// TwinCAT 3 PLC project Untitled1
// ProgramVersion: 3.1.4026.27
// libraries:
//   Tc2_Standard, * (Beckhoff Automation GmbH)
//   Tc2_System, * (Beckhoff Automation GmbH)
//   Tc3_EventLogger, * (Beckhoff Automation GmbH)
//   Tc3_Module, * (Beckhoff Automation GmbH)
//   VisuDialogs, * (System)
//   VisuSymbols,4.5.0.0,System
// project tree:
//   / GlobalTextList.TcGTLO, PlcTask.TcTTO, Visualization Manager.TcVMO (not stored)
//   GVLs/ gAL.TcGVL
//   POUs/Alarms_and_Emergency/ Alarm_System.TcPOU, FB_Emergency_Shutdown.TcPOU, FB_Alarm.TcPOU
//   POUs/ FB_ControlPanel.TcPOU, FB_Scale.TcPOU, MAIN.TcPOU, PI_Function_Block.TcPOU
// real-time tasks:
//   TASK PlcTask: cycle T#10ms, priority 20, ADS port 350
// I/O:
//   DEVICE Device 1 (EtherCAT), AmsNetId 10.0.0.14.2.1
//     Term 7 (EK1200) [EK1200-5000 EtherCAT Power supply (2A E-Bus)]
//       Term 2 (EL4004) [EL4004 4Ch. Ana. Output 0-10V, 12bit]
//       Term 3 (EL4004) [EL4004 4Ch. Ana. Output 0-10V, 12bit]
//       Term 8 (EL3024) [EL3024 4Ch. Ana. Input 4-20mA DIFF]
//       Term 9 (EL3024) [EL3024 4Ch. Ana. Input 4-20mA DIFF]
//       Term 12 (EL1859) [EL1859 8Ch. Dig. Input 24V, 3ms, 8Ch. Dig. Output 24V, 0.5A]
//       Term 13 (EL9011) [EL9011 End Terminal]
//   DEVICE Device 4 (COM Port) (disabled)
// variable links:
//   Untitled1/Untitled1 Instance <-> Device 1 (EtherCAT)/Term 7 (EK1200)/Term 12 (EL1859)
//     PlcTask Inputs/MAIN.EMERGENCY_STOP <-> Channel 1/EMERGENCY STOP
//     PlcTask Inputs/MAIN.Start_Button <-> Channel 2/Start Button
//     PlcTask Inputs/MAIN.Stop_Button <-> Channel 3/Stop Button
//     PlcTask Outputs/MAIN.Motor_Direction <-> Channel 10/Motor Direction
//     PlcTask Outputs/MAIN.Motor_ON_OFF <-> Channel 9/Motor ON/OFF
//   Untitled1/Untitled1 Instance <-> Device 1 (EtherCAT)/Term 7 (EK1200)/Term 2 (EL4004)
//     PlcTask Outputs/MAIN.Flow_Valve_1 <-> AO Outputs Channel 4/Flow_Valve_1
//     PlcTask Outputs/MAIN.Level_Valve_1 <-> AO Outputs Channel 1/Level_Valve_1
//     PlcTask Outputs/MAIN.Level_Valve_2 <-> AO Outputs Channel 2/Level_Valve_2
//     PlcTask Outputs/MAIN.Level_Valve_3 <-> AO Outputs Channel 3/Level_Valve_3
//   Untitled1/Untitled1 Instance <-> Device 1 (EtherCAT)/Term 7 (EK1200)/Term 3 (EL4004)
//     PlcTask Outputs/MAIN.Gas_Valve <-> AO Outputs Channel 1/Gas_Valve
//     PlcTask Outputs/MAIN.Mixer_Valve <-> AO Outputs Channel 2/Mixer_Valve
//     PlcTask Outputs/MAIN.Motor_speed <-> AO Outputs Channel 3/Motor_Speed
//   Untitled1/Untitled1 Instance <-> Device 1 (EtherCAT)/Term 7 (EK1200)/Term 8 (EL3024)
//     PlcTask Inputs/MAIN.Pressure_Differencial_Transmitter_1 <-> AI Standard Channel 1/PDT 1
//     PlcTask Inputs/MAIN.Pressure_Differencial_Transmitter_2 <-> AI Standard Channel 3/PDT 2
//     PlcTask Inputs/MAIN.Pressure_Transmitter_1 <-> AI Standard Channel 2/PT 1
//     PlcTask Inputs/MAIN.Pressure_Transmitter_3 <-> AI Standard Channel 4/PT 3
//   Untitled1/Untitled1 Instance <-> Device 1 (EtherCAT)/Term 7 (EK1200)/Term 9 (EL3024)
//     PlcTask Inputs/MAIN.Level_Transmitter_1 <-> AI Standard Channel 2/ Level Transmitter 1
//     PlcTask Inputs/MAIN.Level_Transmitter_2 <-> AI Standard Channel 3/Level Transmitter 2
//     PlcTask Inputs/MAIN.Pressure_Transmitter_2 <-> AI Standard Channel 1/PT 2
//     PlcTask Inputs/MAIN.Temperature_Transmitter <-> AI Standard Channel 4/Temperature Transmitter

CONFIGURATION Untitled1
    RESOURCE PLC ON TwinCAT3
        TASK PlcTask(INTERVAL := T#10ms, PRIORITY := 20);
        PROGRAM MAIN WITH PlcTask : MAIN;
        PROGRAM Alarm_System WITH PlcTask : Alarm_System;
    END_RESOURCE
END_CONFIGURATION

// ---- GVLs/gAL.TcGVL
{attribute 'qualified_only'}
VAR_GLOBAL
    fbTempWarning  : FB_TcAlarm;
	fbPressWarning : FB_TcAlarm;
	fbTempTrip     : FB_TcAlarm;
	fbPressTrip    : FB_TcAlarm;
	fbEstop        : FB_TcAlarm;
END_VAR

// ---- POUs/MAIN.TcPOU
PROGRAM MAIN
VAR
	//Linking variables to IO cards
	Flow_Valve_1 AT %Q* : INT;
	Level_Valve_1 AT %Q* : INT;
	Level_Valve_2 AT %Q* : INT;
	Level_Valve_3 AT %Q* : INT;
	Gas_Valve AT %Q* : INT;
	Mixer_Valve AT %Q* : INT;
	Motor_speed AT %Q* : INT;
	Motor_ON_OFF AT %Q* :BOOL;
	Motor_Direction AT %Q* :BOOL; 
	Start_Button AT %I* :BOOL;
	Stop_Button AT %I* : BOOL; 
	EMERGENCY_STOP AT %I* : BOOL; 
	Level_Transmitter_1 AT %I* :INT; 
	Level_Transmitter_2 AT %I* :INT; 
	Temperature_Transmitter AT %I* :INT;  
	Pressure_Differencial_Transmitter_1 AT %I* : INT;
	Pressure_Differencial_Transmitter_2 AT %I* : INT;
	Pressure_Transmitter_1 AT %I* : INT ; 
	Pressure_Transmitter_2 AT %I* : INT ; 
	Pressure_Transmitter_3 AT %I* : INT ;
	bSimulate : BOOL := FALSE;   // TRUE = kjører lokalt uten I/O. SETT FALSE PÅ EKTE PLC!
	bReset : BOOL;   // Felles reset fra HMI: alarmer, safe state og motor - olavr

	
	//User Input as percentage
	Flow_Valve_1_Percentage: INT :=100;
	Level_Valve_1_Percentage: INT  := 0;
	Level_Valve_2_Percentage: INT := 0;
	Level_Valve_3_Percentage: INT := 0;
	Motor_speed_Percentage: INT := 0;
	Motor_ON : BOOL ;
	ON_OFF : STRING(10) := 'OFF' ; 
	
	//Scaled values
	Level_Transmitter_1_Scaled : REAL;
	Level_Transmitter_2_Scaled : REAL;
	Pressure_Differential_Transmitter_1_Scaled : REAL;
	Pressure_Differential_Transmitter_2_Scaled : REAL;
	
	//PI function block instantiation
	PI_Controller : PI_Function_Block;
	
	//PI controller on/off state
	bControllerActive : BOOL;
	

    Scale_PT1 : FB_Scale;
	Scale_PT2 : FB_Scale;
	Scale_PT3 : FB_Scale;
	Scale_PDT1: FB_Scale;
	Scale_PDT2: FB_Scale;
    Scale_TT1 : FB_Scale;
	Scale_LT1 : FB_Scale;
	Scale_LT2 : FB_Scale;
    
    Pressure_1_Bar_Scaled : REAL;
	Pressure_2_Bar_Scaled : REAL;
	Pressure_3_Bar_Scaled : REAL;
    Temperature_1_Scaled  : REAL;

	

    bAlarmReset    : BOOL;      // Reset-knapp fra HMI

	fbTempAlarm    : FB_Alarm; // FB_Alarm er røykvarsler-modellen, altså tegningen av hvordan den virker.
	fbPressAlarm   : FB_Alarm;   // fbTempAlarm og fbPressAlarm er to faktiske røykvarslere montert i hvert sitt rom.
	

	// Synlighet for varseltrekant i HMI (trip eller nødstopp) - Variabelen er en string siden HMI
	// Kreven tekst
	
	
	fbEmergency_Shutdown : FB_Emergency_Shutdown;
	
	
	
	// FYSISKE KNAPPER
	fbControlPanel : FB_ControlPanel;
	bHmiStart      : BOOL;
	bHmiStop       : BOOL;
	bHmiEStop      : BOOL;
	
END_VAR

bReset := bAlarmReset OR (Start_Button AND fbEmergency_Shutdown.bTrip);

fbControlPanel(
	bStartPB  := Start_Button,
	bStopPB   := Stop_Button OR bSimulate,
	bEStopPB  := EMERGENCY_STOP OR bSimulate,
	bHmiStart := bHmiStart,
	bHmiStop  := bHmiStop OR fbEmergency_Shutdown.bTrip,
	bHmiEStop := bHmiEStop,
	bReset    := bReset);

// skalerer, regulerer og sender ut signaler

Scale_LT1(RawValue := Level_Transmitter_1, 
          PhysMin := 20.0, 
          PhysMax := 20.5, 
          ScaledValue => Level_Transmitter_1_Scaled);

Scale_LT2(RawValue := Level_Transmitter_2, 
          PhysMin := 50.0, 
          PhysMax := 50.5, 
          ScaledValue => Level_Transmitter_2_Scaled);
		  
// Oppgitt i prosent, fordi de reelle verdiene ikke er kjent.
Scale_PDT1(RawValue := Pressure_Differencial_Transmitter_1, 
          PhysMin := 0.0, 
          PhysMax := 100.0, 
          ScaledValue => Pressure_Differential_Transmitter_1_Scaled);
		  
Scale_PDT2(RawValue := Pressure_Differencial_Transmitter_2, 
          PhysMin := 45.0, 
          PhysMax := 45.5, 
          ScaledValue => Pressure_Differential_Transmitter_2_Scaled);

// Skaler PT1 (f.eks. 0 til 6 bar)
Scale_PT1(RawValue := Pressure_Transmitter_1, 
          PhysMin := 0.0, 
          PhysMax := 6.0, 
          ScaledValue => Pressure_1_Bar_Scaled);
		  
Scale_PT2(RawValue := Pressure_Transmitter_2, 
          PhysMin := 0.0, 
          PhysMax := 6.0, 
          ScaledValue => Pressure_2_Bar_Scaled);
		  
Scale_PT3(RawValue := Pressure_Transmitter_3, 
          PhysMin := 0.0, 
          PhysMax := 6.0, 
          ScaledValue => Pressure_3_Bar_Scaled);

// Skaler TT1 (f.eks. -200 til 850 grader)
Scale_TT1(RawValue := Temperature_Transmitter, 
          PhysMin := -200.0, 
          PhysMax := 850.0, 
          ScaledValue => Temperature_1_Scaled);
		  
// PI-Controller
PI_Controller(Actual := Level_Transmitter_2_scaled,
bEnable := bControllerActive);
Level_Valve_2_Percentage := REAL_TO_INT(PI_Controller.Output);


// variable interval for Flow_Valve_1_Percentage  form 0 to 100  
IF Flow_Valve_1_Percentage > 100 THEN
	Flow_Valve_1_Percentage := 100; 
	ELSE IF Flow_Valve_1_Percentage < 0 THEN 
		Flow_Valve_1_Percentage := 0; 
	END_IF
	
END_IF

// variable interval for Level_Valve_1_Percentage  form 0 to 100  
IF Level_Valve_1_Percentage > 100 THEN
	Level_Valve_1_Percentage := 100; 
	ELSE IF Level_Valve_1_Percentage < 0 THEN 
		Level_Valve_1_Percentage := 0; 
	END_IF
	
END_IF

// variable interval for Level_Valve_2_Percentage  form 0 to 100 
IF Level_Valve_2_Percentage > 100 THEN
	Level_Valve_2_Percentage := 100; 
	ELSE IF Level_Valve_2_Percentage < 0 THEN 
		Level_Valve_2_Percentage := 0; 
	END_IF
	
END_IF

// variable interval for Level_Valve_3_Percentage  form 0 to 100 
IF Level_Valve_3_Percentage > 100 THEN
	Level_Valve_3_Percentage := 100; 
	ELSE IF Level_Valve_3_Percentage < 0 THEN 
		Level_Valve_3_Percentage := 0; 
	END_IF
	
END_IF



// variable interval for Motor_speed_Percentage  form 0 to 100 
IF Motor_speed_Percentage > 100 THEN
	Motor_speed_Percentage := 100; 
	ELSE IF Motor_speed_Percentage < 0 THEN 
		Motor_speed_Percentage := 0; 
	END_IF
	
END_IF

// Motor går når prosessen kjører. Nødstopp/trip håndteres i fbEmergency_Shutdown
Motor_ON_OFF := fbControlPanel.bRunning;

// Flow_Valve_1 calibration
Flow_Valve_1 := REAL_TO_INT (262.14*Flow_Valve_1_Percentage +6553 ); 

// Level_Valve_1 calibration
Level_Valve_1 := REAL_TO_INT(262.14*Level_Valve_1_Percentage +6553);

// Level_Valve_2 calibration
Level_Valve_2 := REAL_TO_INT(262.14*Level_Valve_2_Percentage +6553);

// Level_Valve_3 calibration
Level_Valve_3 := REAL_TO_INT(262.14*Level_Valve_3_Percentage +6553);


// Motor_speed calibration
Motor_speed := REAL_TO_INT(262.14*Motor_speed_Percentage +6553);


fbTempAlarm(rValue := Temperature_1_Scaled, rLimit := 80.0, bReset := bReset);
fbPressAlarm(rValue := MAX(Pressure_1_Bar_Scaled, MAX(Pressure_2_Bar_Scaled, Pressure_3_Bar_Scaled)), rLimit := 4.0, bReset := bReset);

// Alarmhåndtering: sender warnings og trips til EventLogger/HMI
Alarm_System();

	
// Safe state
fbEmergency_Shutdown(
	Motor_ON_OFF      := Motor_ON_OFF,
	bControllerActive := bControllerActive,
	Motor_speed       := Motor_speed,
	Gas_Valve         := Gas_Valve,
	Flow_Valve_1      := Flow_Valve_1,
	Level_Valve_1     := Level_Valve_1,
	Level_Valve_2     := Level_Valve_2,
	Level_Valve_3     := Level_Valve_3);

// Motorstatus til HMI (etter safe state, så den viser riktig)
IF Motor_ON_OFF THEN
	Motor_ON := FALSE;
	ON_OFF   := 'MOTOR: ON';
ELSE
	Motor_ON := TRUE;
	ON_OFF   := 'MOTOR: OFF';
END_IF

END_PROGRAM

// ---- POUs/PI_Function_Block.TcPOU
FUNCTION_BLOCK PI_Function_Block
VAR_INPUT
    Setpoint :REAL := 54;
    Actual: REAL;
	Bias: REAL := 40;
    Kp :REAL := 20;
    Ti :REAL := 40;
    Td :REAL := 0;
    Ts :REAL := 0.01;
    N :REAL := 1;
    OutMax :REAL := 100;
    OutMin :REAL := 0;
    bEuler :BOOL := FALSE;
	bEnable :BOOL;
END_VAR

VAR_OUTPUT
    Output :REAL;
    Error :REAL;
END_VAR

VAR
    PrevError :REAL;
    Integ :REAL;
    Deriv :REAL;
    dInteg :REAL;
    Tf :REAL;
    DerivRaw :REAL;
    Unsat :REAL;
END_VAR

Error := Actual - Setpoint;

IF NOT bEnable THEN
	Integ := 0.0;
	dInteg := 0.0;
	Output := Main.Level_Valve_2_Percentage;
	RETURN;
END_IF

IF Ti > 0.0 THEN
    IF bEuler THEN
    dInteg := Ts / Ti * Error;
ELSE
    dInteg := Ts / Ti * (Error + PrevError) / 2;
END_IF
ELSE
    dInteg := 0.0;
    Integ := 0.0;
END_IF

IF N > 0.0 THEN
    Tf := Td / N;
ELSE
    Tf := 0.0;
END_IF

DerivRaw := Td * (Error - PrevError) / Ts;
Deriv := (Tf * Deriv + Ts * DerivRaw)
/ (Tf + Ts);

Unsat := Kp * (Error + Integ + dInteg + Deriv) + Bias;

IF (Unsat > OutMax AND dInteg > 0) OR
(Unsat < OutMin AND dInteg < 0) THEN
dInteg := 0; // anti-windup
END_IF
Integ := Integ + dInteg;

Output := Kp * (Error + Integ + Deriv) + Bias;
IF Output > OutMax THEN Output := OutMax; END_IF
IF Output < OutMin THEN Output := OutMin; END_IF

PrevError := Error;

END_FUNCTION_BLOCK

// ---- POUs/FB_Scale.TcPOU
FUNCTION_BLOCK FB_Scale
VAR_INPUT
    RawValue : INT;       
    RawMin   : REAL := 0.0;     
    RawMax   : REAL := 32767.0; 
    PhysMin  : REAL;      
    PhysMax  : REAL;      
END_VAR

VAR_OUTPUT
    ScaledValue : REAL;   
END_VAR

// Error handling to prevent division by zero.
IF (RawMax - RawMin) <> 0.0 THEN
    ScaledValue :=  PhysMin + (PhysMax - PhysMin) * (INT_TO_REAL(RawValue) - RawMin) / (RawMax - RawMin);
ELSE
    ScaledValue := PhysMin;
END_IF

END_FUNCTION_BLOCK

// ---- POUs/Alarms_and_Emergency/FB_Alarm.TcPOU
FUNCTION_BLOCK FB_Alarm
VAR_INPUT
	rValue : REAL; // Målt verdi 
	rLimit : REAL; // Maks verdi for BAR og temperatur
	bReset : BOOL; // Denne nulstiller alarmen, denne blir brukt i HMIen
END_VAR
VAR_OUTPUT
	bAlarm  : BOOL;    // TRUE når alarmen er aktiv
END_VAR
VAR
	fbLatch : RS; // Fungerer som minnebryter - Eks: Trykket går under 4 Bar, men alarmen fortsetter å gå, fordi den husker at noe skjedde.
	               // Først når noen trykker reset, slår den seg av.
				   // Det er nettopp det RS gjør. SET slår den på, den blir stående på, og RESET slår den av.
				   // fbLatch er ikke en verdi, men en instans av RS-blokken, altså en egen liten “minnebryter” som lever inne i FB_Alarm
END_VAR

// FB_Alarm er røykvarsleren. Den merker brannen og fortsetter å pipe til noen kvitterer.

//FB_Alarm bestemmer om det er alarm.

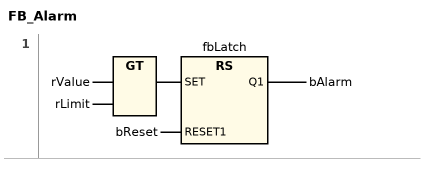
// NETWORK 1
fbLatch(SET := rValue > rLimit, RESET1 := bReset); // RS
bAlarm := fbLatch.Q1;

END_FUNCTION_BLOCK

// ---- POUs/Alarms_and_Emergency/FB_Emergency_Shutdown.TcPOU
FUNCTION_BLOCK FB_Emergency_Shutdown
VAR_INPUT
END_VAR
VAR_OUTPUT
	bTrip : BOOL;          // TRUE = systemet skal stoppes
END_VAR
VAR_IN_OUT
	Motor_ON_OFF      : BOOL;
	bControllerActive : BOOL;
	Motor_speed       : INT;
	Gas_Valve         : INT;
	Flow_Valve_1      : INT;
	Level_Valve_1     : INT;
	Level_Valve_2     : INT;
	Level_Valve_3     : INT;
END_VAR

//MAIN . fbPressAlarm . bAlarm
 //│          │           │
// │          │           └─ variabelen bAlarm inne i den blokken
// │          └─ instansen fbPressAlarm, som er deklarert i MAIN
// └─ programmet MAIN

//Instans: typen er en funksjonsblokk. Den holder en hel pakke, med innganger, utganger og internt minne, og den har kode som kan kjøres.

// Gas_Valve := REAL_TO_INT(262.14 * Prosent + 6553);

// Setter maskinen i safe state
VAR
	fbTripLatch: SR;
END_VAR
VAR // added by the converter: edge detectors and wires of the graphical bodies
    _w1 : BOOL;
END_VAR

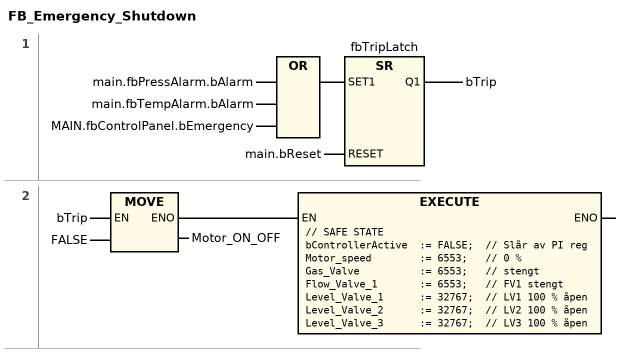
// NETWORK 1
fbTripLatch(SET1 := main.fbPressAlarm.bAlarm OR main.fbTempAlarm.bAlarm OR MAIN.fbControlPanel.bEmergency, RESET := main.bReset); // SR
bTrip := fbTripLatch.Q1;

// NETWORK 2
_w1 := bTrip;
IF _w1 THEN Motor_ON_OFF := FALSE; END_IF
IF _w1 THEN
    // SAFE STATE
    bControllerActive  := FALSE;  // Slår av PI reg 
    Motor_speed        := 6553;   // 0 %
    Gas_Valve          := 6553;   // stengt
    Flow_Valve_1       := 6553;   // FV1 stengt
    Level_Valve_1      := 32767;  // LV1 100 % åpen
    Level_Valve_2      := 32767;  // LV2 100 % åpen
    Level_Valve_3      := 32767;  // LV3 100 % åpen
END_IF

END_FUNCTION_BLOCK

// ---- POUs/FB_ControlPanel.TcPOU
FUNCTION_BLOCK FB_ControlPanel
VAR_INPUT
	bStartPB    : BOOL;  // physical start, NO (TRUE = pressed)
	bStopPB     : BOOL;  // physical stop, NC (FALSE = pressed)
	bEStopPB    : BOOL;  // physical emergency, NC (FALSE = pressed)
	bHmiStart   : BOOL;  // soft buttons from HMI
	bHmiStop    : BOOL;
	bHmiEStop   : BOOL;
	bReset      : BOOL;  // felles reset (HMI)
END_VAR
VAR_OUTPUT
	bRunning    : BOOL;  // process is allowed to run
	bEmergency  : BOOL;  // latched emergency, needs reset
	bStopActive : BOOL;  // a stop is being requested right now
END_VAR
VAR
	rtStart     : R_TRIG;
	rtHmiStart  : R_TRIG;
END_VAR

// Flankedeteksjon på start
rtStart(CLK := bStartPB);
rtHmiStart(CLK := bHmiStart);

// Stopp = fysisk NC åpnet ELLER soft stop (inkl. trip fra MAIN)
bStopActive := NOT bStopPB OR bHmiStop;

// Nødstopp låses. Kvitteres kun med bReset når nødstoppen er sluppet
IF NOT bEStopPB OR bHmiEStop THEN
	bEmergency := TRUE;
ELSIF bEmergency AND bReset THEN
	bEmergency := FALSE;
END_IF

// Start på stigende flanke, kun når ingen stopp eller nødstopp er aktiv
IF bEmergency OR bStopActive THEN
	bRunning := FALSE;
ELSIF rtStart.Q OR rtHmiStart.Q THEN
	bRunning := TRUE;
END_IF

END_FUNCTION_BLOCK

// ---- POUs/Alarms_and_Emergency/Alarm_System.TcPOU
PROGRAM Alarm_System
VAR
	bAlarmsCreated : BOOL;
END_VAR


// Alarm_System er alarmsentralen. Den logger og viser alarmen i HMI-en.

// Alarm_System melder fra om alarmen.

// Opprett alarmene én gang ved oppstart
// 2. param: FALSE = warning (forsvinner selv), TRUE = trip/nødstopp (må kvitteres)
IF NOT bAlarmsCreated THEN
    bAlarmsCreated := TRUE;
    gAL.fbTempWarning.CreateEx(TC_EVENTS.ProcessAlarmEvent.HighTemperatureWarning, FALSE, 0);
    gAL.fbPressWarning.CreateEx(TC_EVENTS.ProcessAlarmEvent.HighPressureWarning, FALSE, 0);
    gAL.fbTempTrip.CreateEx(TC_EVENTS.ProcessAlarmEvent.HighTemperature, TRUE, 0);
    gAL.fbPressTrip.CreateEx(TC_EVENTS.ProcessAlarmEvent.HighPressure, TRUE, 0);
    gAL.fbEstop.CreateEx(TC_EVENTS.ProcessAlarmEvent.EmergencyButtonPressed, TRUE, 0);
END_IF

// Warnings: aktive så lenge verdien er over grensen
IF MAIN.Temperature_1_Scaled > 70.0 THEN
    IF NOT gAL.fbTempWarning.bRaised THEN gAL.fbTempWarning.Raise(0); END_IF
ELSIF gAL.fbTempWarning.bRaised THEN
    gAL.fbTempWarning.Clear(0, FALSE);
END_IF

IF MAIN.Pressure_1_Bar_Scaled > 3.5 THEN
    IF NOT gAL.fbPressWarning.bRaised THEN gAL.fbPressWarning.Raise(0); END_IF
ELSIF gAL.fbPressWarning.bRaised THEN
    gAL.fbPressWarning.Clear(0, FALSE);
END_IF

// Trips: følger FB_Alarm i MAIN (låst til Reset)
IF MAIN.fbTempAlarm.bAlarm THEN
    IF NOT gAL.fbTempTrip.bRaised THEN gAL.fbTempTrip.Raise(0); END_IF
ELSIF gAL.fbTempTrip.bRaised THEN
    gAL.fbTempTrip.Clear(0, FALSE);
END_IF

IF MAIN.fbPressAlarm.bAlarm THEN
    IF NOT gAL.fbPressTrip.bRaised THEN gAL.fbPressTrip.Raise(0); END_IF
ELSIF gAL.fbPressTrip.bRaised THEN
    gAL.fbPressTrip.Clear(0, FALSE);
END_IF

// Nødstopp
IF MAIN.fbControlPanel.bEmergency THEN
    IF NOT gAL.fbEstop.bRaised THEN gAL.fbEstop.Raise(0); END_IF
ELSIF gAL.fbEstop.bRaised THEN
    gAL.fbEstop.Clear(0, FALSE);
END_IF

END_PROGRAM

// ---- GlobalTextList.TcGTLO
TEXTLIST GlobalTextList
  9 = '%f'
  594 = '%I'
  907 = '%i'
  617 = 'aaaaaaaa'
  411 = 'EMERGENCY STOP'
  749 = 'EMERGENCY STOP %s'
  283 = 'Flow Valve %i'
  422 = 'Flow Valve 1 = %f %'
  201 = 'Flow Valve = %i'
  842 = 'Flow Valve: %i'
  336 = 'Flow Valve: %i %'
  590 = 'Flow Valve: %i%'
  567 = 'Gas Valve : %i%'
  736 = 'Level Valve 1 = %f %'
  833 = 'Level Valve 1 = %i %'
  36 = 'Level Valve 1: %i'
  942 = 'Level Valve 1: %i%'
  802 = 'Level Valve 2: %i%'
  940 = 'Level Valve 3: %i%'
  781 = 'Mixer Valve : %i%'
  1 = 'Motor   %s'
  109 = 'Motor Direction %s'
  202 = 'Motor OFF'
  60 = 'Motor OFF  '
  480 = 'Motor OFF  %B'
  834 = 'Motor OFF  %s'
  840 = 'Motor ON'
  885 = 'MOtor ON'
  981 = 'Motor Speed: %i%'
  390 = 'PDT 1'
  74 = 'PDT 1 %i'
  240 = 'PDT 1 = %.4f  Bar'
  2 = 'PDT 1 = %4.f  Bar'
  419 = 'PDT 1 = %4f  Bar'
  414 = 'PDT 1 = %f Bar'
  882 = 'PDT 1 = %f.4 Bar'
  541 = 'PDT 1 = %fmaxDecimals = 3 Bar'
  384 = 'PDT 1 = %i'
  145 = 'PDT 1 = %i Bar'
  423 = 'PDT 2 %i'
  214 = 'PDT 2 = %.4f Bar'
  437 = 'PDT 2 = %f Bar'
  723 = 'PDT 2 = %i'
  493 = 'PDT 2 = %i Bar'
  589 = 'PT 1 %i'
  999 = 'PT 1 = %.4f Bar'
  314 = 'PT 1 = %f Bar'
  203 = 'PT 1 = %i Bar'
  730 = 'sdfsdf'
  313 = 'START'
  187 = 'START %s'
  945 = 'STOP'
  921 = 'STOP %s'
END_TEXTLIST
